{region 'Documentation'}
(*!
<summary>Check that IN is strictly later than Minimum.</summary>
*)
{endregion}
FUNCTION_BLOCK AssertLaterThan_LTime EXTENDS AssertionBase
VAR_INPUT
    IN : LTIME; //! Actual value checked or observed by this Assertion.
    Minimum : LTIME; //! Exclusive lower bound; the actual value or count must be greater.
END_VAR

SUPER^();

{region 'Documentation'}
(*!
<summary>Evaluate the typed duration relation and report higher-priority errors first.</summary>
*)
{endregion}
METHOD PROTECTED Assert
VAR
    Message : STRING(GVL_Constants.MessageLength);
    MinimumText : STRING(GVL_Constants.AssertionValueLength);
    ActualText : STRING(GVL_Constants.AssertionValueLength);
END_VAR
IF NOT EvaluationActive THEN
    RETURN;
END_IF;

IF Result = E_Result.Error THEN
    RETURN;
END_IF;

IF Result = E_Result.Failed THEN
    RETURN;
END_IF;

IF IN <= Minimum THEN
    MinimumText := LTIME_TO_STRING(Minimum);
    ActualText := LTIME_TO_STRING(IN);
    Message := CONCAT('Assertion failed: value is not later than limit. Minimum = ',
        MinimumText);
    Message := CONCAT(Message, ', Actual = ');
    Message := CONCAT(Message, ActualText);
    Message := CONCAT(Message, '.');
    Fail(Message := Message);
    RETURN;
END_IF;

Pass();
END_METHOD

END_FUNCTION_BLOCK

(* stored: Version 1.1.0.1
   POU AssertLaterThan_LTime: Id {f9d33c42-9dcf-4632-9259-235b9a84ebe9}, SpecialFunc None
   Folder Internal: Id {b9175fa3-bf9e-4bd4-bf7d-67e3d82ca659}
   Method Assert: Id {5349a671-8158-43da-8145-ce6d9e0aedae} *)
